Fanuc KAREL source: kx00010.KL

-- PROVISIONAL review KL for V1013-1; original PC SHA256 56cb0805213124cf52772c720b131cb00d79eddcc41d56f7b64fb2a330ab3b78
-- Incomplete behavior may be omitted. Consult companion uncertainty JSON. Do not deploy.
PROGRAM KX00010
%NOLOCKGROUP
VAR
  I : INTEGER
  J : INTEGER
  B : BOOLEAN
  F : FILE
  S : STRING[80]
-- UNRESOLVED_DECL P type=000102
BEGIN
  -- UNRESOLVED_PC offsets 5-7; opcodes 9C,10
  -- UNRESOLVED_PC offsets 12-16; opcodes 7F
END KX00010
